(* IEC 61131-3 sources: BODAS-RC27-18_40/st/bodas_rc18_12_27_18_40/plc_logic/application/easyconfig_import/bdl, 8 files *)

(* ---- bds_snsrdsa_inst_te-bds_snsrDsa_inst_te.st ---- *)
(* --- Interface --- *)
{attribute 'qualified_only' := ''}
{attribute 'strict' := ''}
TYPE bds_snsrDsa_inst_te :
(
	bds_snsrDsa_numInst_E := 0
) USINT;
END_TYPE

(* ---- bds_snsrdsa_inst_te_1-bds_snsrDsa_inst_te_1.st ---- *)
(* --- Interface --- *)
{attribute 'qualified_only' := ''}
{attribute 'strict' := ''}
TYPE bds_snsrDsa_inst_te_1 :
(
	bds_snsrDsa_numInst_E
) USINT;
END_TYPE

(* ---- bds_snsrdst_inst_te-bds_snsrDst_inst_te.st ---- *)
(* --- Interface --- *)
{attribute 'qualified_only' := ''}
{attribute 'strict' := ''}
TYPE bds_snsrDst_inst_te :
(
	bds_snsrDst_numInst_E
) USINT;
END_TYPE

(* ---- bds_snsrdst_inst_te_1-bds_snsrDst_inst_te_1.st ---- *)
(* --- Interface --- *)
{attribute 'qualified_only' := ''}
{attribute 'strict' := ''}
TYPE bds_snsrDst_inst_te_1 :
(
	bds_snsrDst_numInst_E
) USINT;
END_TYPE

(* ---- bds_snsrpal_inst_te-bds_snsrPal_inst_te.st ---- *)
(* --- Interface --- *)
{attribute 'qualified_only' := ''}
{attribute 'strict' := ''}
TYPE bds_snsrPal_inst_te :
(
	bds_snsrPal_numInst_E := 0
) USINT;
END_TYPE

(* ---- bds_snsrpal_inst_te_1-bds_snsrPal_inst_te_1.st ---- *)
(* --- Interface --- *)
{attribute 'qualified_only' := ''}
{attribute 'strict' := ''}
TYPE bds_snsrPal_inst_te_1 :
(
	bds_snsrPal_numInst_E
) USINT;
END_TYPE

(* ---- bds_snsrpr4_inst_te-bds_snsrPr4_inst_te.st ---- *)
(* --- Interface --- *)
{attribute 'qualified_only' := ''}
{attribute 'strict' := ''}
TYPE bds_snsrPr4_inst_te :
(
	bds_snsrPr4_numInst_E := 0
) USINT;
END_TYPE

(* ---- bds_snsrpr4_inst_te_1-bds_snsrPr4_inst_te_1.st ---- *)
(* --- Interface --- *)
{attribute 'qualified_only' := ''}
{attribute 'strict' := ''}
TYPE bds_snsrPr4_inst_te_1 :
(
	bds_snsrPr4_numInst_E := 0
) USINT;
END_TYPE
